// TIA Portal V20 export
FUNCTION "Zählerfunktion mit STOP" : Void   // FC106, STL
TITLE = Zählerfunktion mit Stop
{ S7_Optimized_Access := 'FALSE' }
AUTHOR : SD
FAMILY : Zähler
// stored: AutoNumber false
   VAR_INPUT
      Stopwert : DInt;   // Bei diesem Wert wird ein Stopsignal ausgegeben
      RESET : Bool;
   END_VAR
   VAR_IN_OUT
      Zaehlsignal : Bool;
      Zaehlerstand : DInt;
      Stopbit : Bool;   // Stopbit
   END_VAR
BEGIN

NETWORK
TITLE = Zählsignal
      AN    #Zaehlsignal;
      JC    M031;

      SET;
      R     #Zaehlsignal;

NETWORK
TITLE = Zählerstand erhöhen
      L     #Zaehlerstand;
      L     1;
      +D;
      T     #Zaehlerstand;

NETWORK
TITLE = Vergleich von Ist und Sollstand
      L     #Zaehlerstand;
      L     #Stopwert;
      <D;
      JC    M031;
      SET;
      S     #Stopbit;

M031: NOP   0;

NETWORK
TITLE = Reset Stopbit und Zählerstand
      AN    #RESET;
      JC    M041;
      L     0;
      T     #Zaehlerstand;

      SET;
      R     #Stopbit;
M041: NOP   0;
END_FUNCTION
